// TIA Portal V21 export
// export: Created 2026-11-11T00:47:19.7091716Z, ExportSetting WithDefaults, DisplayName Totally Integrated Automation Portal, DisplayVersion V21 Update 3, DisplayName STEP 7 Professional, DisplayVersion V21 Update 3, DisplayName STEP 7 Safety, DisplayVersion V21, DisplayName Tech WebApplication, DisplayVersion V21, DisplayName WinCC Basic/Comfort/Advanced, DisplayVersion V21 Update 3, DisplayName WinCC Unified, DisplayVersion V21 Update 3
FUNCTION_BLOCK "FB_Fbd_ex057"   // FB95, FBD
{ S7_Optimized_Access := 'TRUE' }
VERSION : 0.1
// stored: AutoNumber true, IsIECCheckEnabled false, IsRetainMemResEnabled false, MemoryReserve 100, SetENOAutomatically false, UDAEnableTagReadback false
   VAR_INPUT
      v_req : Bool;
      v_mode : UInt;
      v_laddr : HW_INTERFACE;
      v_ctrlrec : Array[0..99] of Byte;
   END_VAR
   VAR_OUTPUT
      v_done : Bool;
      v_busy : Bool;
      v_error : Bool;
      v_status : DWord;
      v_err_info : Word;
   END_VAR
   VAR
      inst { S7_SetPoint := 'True'} : ReconfigIOSystem;
   END_VAR
BEGIN

REGION Network 1: ReconfigIOSystem - Reconfigure IO system
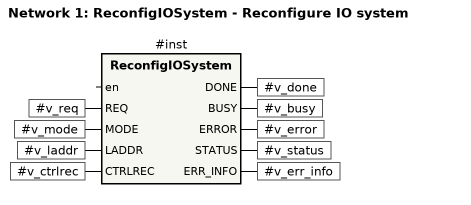
   #inst(REQ := #v_req,   // ReconfigIOSystem
         MODE := #v_mode,
         LADDR := #v_laddr,
         CTRLREC := #v_ctrlrec,
         DONE => #v_done,
         BUSY => #v_busy,
         ERROR => #v_error,
         STATUS => #v_status,
         ERR_INFO => #v_err_info);
END_REGION
END_FUNCTION_BLOCK
